// TIA Portal V21 export
Screen "R06a_MoveH"  1024x768, Number=45, Template=Tpl
  ScreenLayer 
    IOField "P_CraneX" at 10,10 size 100x30  Mode=Output
      ProcessValue := P_Cell
      HorizontalMovementAnimation "HorizontalMovementAnimation"
